(* IEC 61131-3 sources: rusty/tests/lit/single/builtin, 48 files *)

(* ---- abs_arguments.st ---- *)
// RUN: %COMPILE %s && %RUN | %CHECK %s
//
// ABS gives the same result for the implicit (positional) and the explicit (named) call form.

FUNCTION main
VAR
    neg : DINT := -42;
    a   : DINT;
    b   : DINT;
END_VAR

a := ABS(neg);
b := ABS(IN := neg);
// CHECK: ABS=42 42
printf('ABS=%d %d$N', a, b);
END_FUNCTION

(* ---- abs_floats.st ---- *)
// RUN: %COMPILE %s && %RUN | %CHECK %s
//
// ABS on floats lowers to the llvm.fabs intrinsic.

FUNCTION main

// CHECK: real=3.2 0.0 3.3 0.0
printf('real=%.1f %.1f %.1f %.1f$N', ABS(REAL#-3.2), ABS(REAL#-0.0), ABS(REAL#3.3), ABS(REAL#0.0));

// CHECK: lreal=2.5 0.0 2.6 0.0
printf('lreal=%.1f %.1f %.1f %.1f$N', ABS(LREAL#-2.5), ABS(LREAL#-0.0), ABS(LREAL#2.6), ABS(LREAL#0.0));
END_FUNCTION

(* ---- abs_signed.st ---- *)
// RUN: %COMPILE %s && %RUN | %CHECK %s
//
// ABS is a builtin; signed integers lower to the llvm.abs intrinsic with
// is_int_min_poison = false, so ABS(INT_MIN) wraps to INT_MIN.

FUNCTION main
VAR
    min : INT := INT#-32768;
END_VAR

// CHECK: sint=120 0 121 0
printf('sint=%d %d %d %d$N', ABS(SINT#-120), ABS(SINT#-0), ABS(SINT#121), ABS(SINT#0));

// CHECK: int=99 0 98 0
printf('int=%d %d %d %d$N', ABS(INT#-99), ABS(INT#-0), ABS(INT#98), ABS(INT#0));

// CHECK: dint=77 0 78 0
printf('dint=%d %d %d %d$N', ABS(-77), ABS(-0), ABS(78), ABS(0));

// CHECK: lint=88 0 89 0
printf('lint=%lld %lld %lld %lld$N', ABS(LINT#-88), ABS(LINT#-0), ABS(LINT#89), ABS(LINT#0));

// CHECK: big=1234567890123
printf('big=%lld$N', ABS(LINT#-1234567890123));

// CHECK: min=-32768
printf('min=%d$N', ABS(min));

// explicit calls to the library monomorphs still link against the stdlib
// CHECK: lib=7
printf('lib=%d$N', ABS__DINT(DINT#-7));
END_FUNCTION

(* ---- abs_unsigned.st ---- *)
// RUN: %COMPILE %s && %RUN | %CHECK %s
//
// ABS of an unsigned value returns the value unchanged instead of calling a
// non-existent monomorph (previously a crash at runtime). Each call reports
// warning E150, see abs_unsigned_warning.st.

FUNCTION main
VAR
    u8  : USINT := USINT#200;
    u16 : UINT  := UINT#5;
    u32 : UDINT := UDINT#4000000000;
    u64 : ULINT := ULINT#42;
END_VAR

// CHECK: u8=200
printf('u8=%d$N', ABS(u8));

// CHECK: u16=5
printf('u16=%d$N', ABS(u16));

// CHECK: u32=4000000000
printf('u32=%u$N', ABS(u32));

// CHECK: u64=42
printf('u64=%llu$N', ABS(u64));
END_FUNCTION

(* ---- abs_unsigned_warning.st ---- *)
// RUN: %COMPILE %s 2>&1 | %CHECK %s
//
// ABS of an unsigned value has no effect and reports a warning for each call.

FUNCTION main
VAR
    u8  : USINT;
    u16 : UINT;
    u32 : UDINT;
    u64 : ULINT;
    res : ULINT;
END_VAR

// CHECK: {{.*}}warning[E150]{{.*}}ABS on a value of unsigned type 'USINT' has no effect{{.*}}
res := ABS(u8);

// CHECK: {{.*}}warning[E150]{{.*}}ABS on a value of unsigned type 'UINT' has no effect{{.*}}
res := ABS(u16);

// CHECK: {{.*}}warning[E150]{{.*}}ABS on a value of unsigned type 'UDINT' has no effect{{.*}}
res := ABS(u32);

// CHECK: {{.*}}warning[E150]{{.*}}ABS on a value of unsigned type 'ULINT' has no effect{{.*}}
res := ABS(u64);
END_FUNCTION

(* ---- add_arguments.st ---- *)
// RUN: %COMPILE %s && %RUN | %CHECK %s
//
// ADD declares a single variadic parameter. A variadic parameter cannot be named, thus ADD has an
// implicit (positional) call form only. The form is extensible.

FUNCTION main
VAR
    x : DINT := 9;
    y : DINT := 7331;
    z : DINT := 60;
    a : DINT;
    b : DINT;
END_VAR

a := ADD(x, y);
b := ADD(x, y, z);
// CHECK: ADD=7340 7400
printf('ADD=%d %d$N', a, b);
END_FUNCTION

(* ---- add_mul_named_argument.st ---- *)
// RUN: not %COMPILE %s --error-format clang 2>&1 | %CHECK %s
//
// ADD and MUL declare a single variadic parameter, which has no name. A named argument is
// rejected, also IN1 and also with the standard library linked.

FUNCTION main : DINT
VAR
    a : DINT := 1;
    b : DINT := 2;
END_VAR
    // CHECK: {{.*}}add_mul_named_argument.st:[[@LINE+2]]:{{[0-9]+}}:{{.*}}error[E089]: Invalid call parameters
    // CHECK-NEXT: {{.*}}add_mul_named_argument.st:[[@LINE+1]]:{{[0-9]+}}:{{.*}}error[E048]: Could not resolve reference to IN1
    main := ADD(IN1 := a, b);
    // CHECK-NEXT: {{.*}}add_mul_named_argument.st:[[@LINE+2]]:{{[0-9]+}}:{{.*}}error[E089]: Invalid call parameters
    // CHECK-NEXT: {{.*}}add_mul_named_argument.st:[[@LINE+1]]:{{[0-9]+}}:{{.*}}error[E048]: Could not resolve reference to IN1
    main := MUL(IN1 := a, b);
    // CHECK-NEXT: error: Compilation aborted due to critical errors
END_FUNCTION

(* ---- adr_arguments.st ---- *)
// RUN: %COMPILE %s && %RUN | %CHECK %s
//
// ADR returns the same address for the implicit (positional) and the explicit (named) call form.

FUNCTION main
VAR
    i : INT := 5;
    p : BOOL;
END_VAR

p := ADR(i) = ADR(IN := i);
// CHECK: ADR=1
printf('ADR=%d$N', p);
END_FUNCTION

(* ---- adr_ptr_arith_runtime.st ---- *)
// RUN: %COMPILE %s && %RUN | %CHECK %s
//
// `ADR(x) + N` is byte-stride pointer arithmetic — `ADR` is declared to
// return LWORD, so the `+` flows through the integer-arithmetic path; the
// receiver pointer ends up `N` bytes past the operand. Regression for #1749
// (previously panicked in `create_llvm_int_binary_expression`).

FUNCTION main
VAR
    arr : ARRAY[0..7] OF BYTE := [0, 0, 0, 0, 0, 0, 0, 0];
    pt  : REF_TO BYTE;
END_VAR

pt := ADR(arr) + 4;
pt^ := BYTE#16#AB;

// CHECK: arr[4]=171
printf('arr[4]=%d$N', arr[4]);

pt := ADR(arr) + 7;
pt^ := BYTE#16#5C;

// CHECK: arr[7]=92
printf('arr[7]=%d$N', arr[7]);

// Subtraction flows through the same path: take a pointer past the end
// and walk back. Writing to arr[2] via `ADR(arr[6]) - 4`.
pt := ADR(arr[6]) - 4;
pt^ := BYTE#16#11;

// CHECK: arr[2]=17
printf('arr[2]=%d$N', arr[2]);
END_FUNCTION

(* ---- and_arguments.st ---- *)
// RUN: %COMPILE %s && %RUN | %CHECK %s
//
// AND declares a single variadic parameter. A variadic parameter cannot be named, thus AND has an
// implicit (positional) call form only. The form is extensible. AND gives the same result as the
// `AND` operator, for BOOL values as well as for bit and integer values.

FUNCTION main
VAR
    t : BOOL := TRUE;
    f : BOOL := FALSE;
    x : BYTE := 16#F0;
    y : BYTE := 16#3C;
    z : BYTE := 16#18;
    i : DINT := 12;
    j : DINT := 10;
    a : BOOL;
    b : BOOL;
    c : BYTE;
    d : BYTE;
    e : DINT;
END_VAR

a := AND(t, t);
b := AND(t, t, f);
// CHECK: AND=1 0 1 0
printf('AND=%u %u %u %u$N', a, b, t AND t, t AND t AND f);

c := AND(x, y);
d := AND(x, y, z);
e := AND(i, j);
// CHECK: AND-bits=48 16 8
printf('AND-bits=%u %u %d$N', c, d, e);
// CHECK: AND-bits-operator=48 16 8
printf('AND-bits-operator=%u %u %d$N', x AND y, x AND y AND z, i AND j);
END_FUNCTION

(* ---- arithmetic_bit_strings.st ---- *)
// RUN: %COMPILE %s 2> %t.err && %RUN | %CHECK %s
// RUN: not grep -E "error|warning" %t.err
//
// ADD, SUB, MUL and DIV accept bit strings as their operators do, and compute the same values.

FUNCTION main : DINT
VAR
    b : BYTE := 16#FF;
    dw : DWORD := 16#100;
    di : DINT := 7;
END_VAR

// CHECK: ADD BYTE 256 256
printf('ADD BYTE %u %u$N', ADD(b, 1), b + 1);
// CHECK-NEXT: SUB DWORD 255 255
printf('SUB DWORD %u %u$N', SUB(dw, 1), dw - 1);
// CHECK-NEXT: SUB named 255 255
printf('SUB named %u %u$N', SUB(IN2 := 1, IN1 := dw), dw - 1);
// CHECK-NEXT: MUL DWORD 65536 65536
printf('MUL DWORD %u %u$N', MUL(dw, dw), dw * dw);
// CHECK-NEXT: DIV DWORD 128 128
printf('DIV DWORD %u %u$N', DIV(dw, 2), dw / 2);
// CHECK-NEXT: ADD DINT BYTE 262 262
printf('ADD DINT BYTE %d %d$N', ADD(di, b), di + b);
END_FUNCTION

(* ---- datetime_arithmetic_chain.st ---- *)
// RUN: %COMPILE %s && %RUN | %CHECK %s
// Chains of date and time arithmetic, in operator and builtin form

FUNCTION main
    VAR
        x : DT := DT#2027-05-05-22:30:15;
        y : TIME := TIME#20s;
        z : TOD := TOD#23:58:00;
    END_VAR

    x := x + y + y + TIME#2h555s;
    printf('%s$N', REF(DT_TO_STRING(x)));                                           // CHECK: DT#2027-05-06-00:40:10

    z := z + TIME#2m5s;
    printf('%s$N', REF(TOD_TO_STRING(z)));                                          // CHECK: TOD#00:00:05

    x := ADD(x, y, MUL(y, 2));
    printf('%s$N', REF(DT_TO_STRING(x)));                                           // CHECK: DT#2027-05-06-00:41:10

    z := SUB(z, TIME#10s);
    printf('%s$N', REF(TOD_TO_STRING(z)));                                          // CHECK: TOD#23:59:55

END_FUNCTION

(* ---- datetime_arithmetic_date.st ---- *)
// RUN: %COMPILE %s && %RUN | %CHECK %s
// Test DATE arithmetic operations return correct types and values

FUNCTION main
    VAR
        date1 : DATE;
        date2 : DATE;
        result : TIME;
    END_VAR

    // SUB_DATE_DATE: DATE - DATE -> TIME (u32)
    date1 := DATE#2024-01-15;
    date2 := DATE#2024-01-10;
    result := SUB_DATE_DATE(date1, date2);
    printf('%s$N', REF(TIME_TO_STRING(result)));                                    // CHECK: T#5d

    // The operators carry out the same functions
    result := date1 - date2;
    printf('%s$N', REF(TIME_TO_STRING(result)));                                    // CHECK: T#5d

    // The builtins carry out the same functions as the operators
    result := SUB(date1, date2);
    printf('%s$N', REF(TIME_TO_STRING(result)));                                    // CHECK: T#5d

END_FUNCTION

(* ---- datetime_arithmetic_dt.st ---- *)
// RUN: %COMPILE %s && %RUN | %CHECK %s
// Test DT arithmetic operations return correct types and values

FUNCTION main
    VAR
        dt1 : DT;
        dt2 : DT;
        t1 : TIME;
        result : TIME;
        dt_result : DT;
    END_VAR

    // ADD_DT_TIME: DT + TIME -> DT (u32)
    dt1 := DT#2024-01-15-12:30:00;
    t1 := TIME#5s;
    dt_result := ADD_DT_TIME(dt1, t1);
    printf('%s$N', REF(DT_TO_STRING(dt_result)));                                   // CHECK: DT#2024-01-15-12:30:05

    // SUB_DT_TIME: DT - TIME -> DT (u32)
    dt1 := DT#2024-01-15-12:30:05;
    t1 := TIME#3s;
    dt_result := SUB_DT_TIME(dt1, t1);
    printf('%s$N', REF(DT_TO_STRING(dt_result)));                                   // CHECK: DT#2024-01-15-12:30:02

    // SUB_DT_DT: DT - DT -> TIME (u32)
    dt1 := DT#2024-01-15-12:30:10;
    dt2 := DT#2024-01-15-12:30:00;
    result := SUB_DT_DT(dt1, dt2);
    printf('%s$N', REF(TIME_TO_STRING(result)));                                    // CHECK: T#10s

    // The operators carry out the same functions
    dt_result := dt1 + t1;
    printf('%s$N', REF(DT_TO_STRING(dt_result)));                                   // CHECK: DT#2024-01-15-12:30:13
    dt_result := dt1 - t1;
    printf('%s$N', REF(DT_TO_STRING(dt_result)));                                   // CHECK: DT#2024-01-15-12:30:07
    result := dt1 - dt2;
    printf('%s$N', REF(TIME_TO_STRING(result)));                                    // CHECK: T#10s

    // The builtins carry out the same functions as the operators
    dt_result := ADD(dt1, t1, T#1m);
    printf('%s$N', REF(DT_TO_STRING(dt_result)));                                   // CHECK: DT#2024-01-15-12:31:13
    result := SUB(dt1, dt2);
    printf('%s$N', REF(TIME_TO_STRING(result)));                                    // CHECK: T#10s

END_FUNCTION

(* ---- datetime_arithmetic_ldate.st ---- *)
// RUN: %COMPILE %s && %RUN | %CHECK %s
// Test LDATE arithmetic operations return correct types and values

FUNCTION main
    VAR
        ldate1 : LDATE;
        ldate2 : LDATE;
        lresult : LTIME;
    END_VAR

    // SUB_LDATE_LDATE: LDATE - LDATE -> LTIME (i64)
    ldate1 := LDATE#2024-01-15;
    ldate2 := LDATE#2024-01-10;
    lresult := SUB_LDATE_LDATE(ldate1, ldate2);
    printf('%s$N', REF(LTIME_TO_STRING(lresult)));                                  // CHECK: LTIME#5d

    // The operators carry out the same functions
    lresult := ldate1 - ldate2;
    printf('%s$N', REF(LTIME_TO_STRING(lresult)));                                  // CHECK: LTIME#5d

    // The builtins carry out the same functions as the operators
    lresult := SUB(ldate1, ldate2);
    printf('%s$N', REF(LTIME_TO_STRING(lresult)));                                  // CHECK: LTIME#5d

END_FUNCTION

(* ---- datetime_arithmetic_ldt.st ---- *)
// RUN: %COMPILE %s && %RUN | %CHECK %s
// Test LDT arithmetic operations return correct types and values

FUNCTION main
    VAR
        ldt1 : LDT;
        ldt2 : LDT;
        lt1 : LTIME;
        lresult : LTIME;
        ldt_result : LDT;
    END_VAR

    // ADD_LDT_LTIME: LDT + LTIME -> LDT (i64, nanosecond precision)
    ldt1 := LDT#2024-01-15-12:30:00;
    lt1 := LTIME#5s;
    ldt_result := ADD_LDT_LTIME(ldt1, lt1);
    printf('%s$N', REF(LDT_TO_STRING(ldt_result)));                                 // CHECK: LDT#2024-01-15-12:30:05

    // SUB_LDT_LTIME: LDT - LTIME -> LDT (i64)
    ldt1 := LDT#2024-01-15-12:30:05;
    lt1 := LTIME#3s;
    ldt_result := SUB_LDT_LTIME(ldt1, lt1);
    printf('%s$N', REF(LDT_TO_STRING(ldt_result)));                                 // CHECK: LDT#2024-01-15-12:30:02

    // SUB_LDT_LDT: LDT - LDT -> LTIME (i64, result is difference in nanoseconds)
    ldt1 := LDT#2024-01-15-12:30:10;
    ldt2 := LDT#2024-01-15-12:30:00;
    lresult := SUB_LDT_LDT(ldt1, ldt2);
    printf('%s$N', REF(LTIME_TO_STRING(lresult)));                                  // CHECK: LTIME#10s

    // The operators carry out the same functions
    ldt_result := ldt1 + lt1;
    printf('%s$N', REF(LDT_TO_STRING(ldt_result)));                                 // CHECK: LDT#2024-01-15-12:30:13
    ldt_result := ldt1 - lt1;
    printf('%s$N', REF(LDT_TO_STRING(ldt_result)));                                 // CHECK: LDT#2024-01-15-12:30:07
    lresult := ldt1 - ldt2;
    printf('%s$N', REF(LTIME_TO_STRING(lresult)));                                  // CHECK: LTIME#10s

    // The builtins carry out the same functions as the operators
    ldt_result := ADD(ldt1, lt1, lt1);
    printf('%s$N', REF(LDT_TO_STRING(ldt_result)));                                 // CHECK: LDT#2024-01-15-12:30:16
    lresult := SUB(ldt1, ldt2);
    printf('%s$N', REF(LTIME_TO_STRING(lresult)));                                  // CHECK: LTIME#10s

END_FUNCTION

(* ---- datetime_arithmetic_long_chain.st ---- *)
// RUN: %COMPILE %s && %RUN | %CHECK %s
// A long chain of date and time arithmetic compiles in time linear to its length

FUNCTION main
    VAR
        t : TIME := TIME#1s;
    END_VAR

    t := ADD(t, t, t, t, t, t, t, t, t, t, t, t, t, t, t, t, t, t, t, t, t, t, t, t, t, t, t, t, t, t);
    printf('%s$N', REF(TIME_TO_STRING(t)));                                         // CHECK: T#30s

    t := t + t + t + t + t + t + t + t + t + t + t + t + t + t + t + t + t + t + t + t + t + t + t + t + t + t + t + t + t + t;
    printf('%s$N', REF(TIME_TO_STRING(t)));                                         // CHECK: T#15m

END_FUNCTION

(* ---- datetime_arithmetic_ltime.st ---- *)
// RUN: %COMPILE %s && %RUN | %CHECK %s
// Test LTIME arithmetic operations return correct types and values

FUNCTION main
    VAR
        lt1 : LTIME;
        lt2 : LTIME;
        lresult : LTIME;
    END_VAR

    // ADD_LTIME: LTIME + LTIME -> LTIME (i64)
    lt1 := LTIME#5s;
    lt2 := LTIME#3s;
    lresult := ADD_LTIME(lt1, lt2);
    printf('%s$N', REF(LTIME_TO_STRING(lresult)));                                  // CHECK: LTIME#8s

    // SUB_LTIME: LTIME - LTIME -> LTIME (i64)
    lt1 := LTIME#10s;
    lt2 := LTIME#3s;
    lresult := SUB_LTIME(lt1, lt2);
    printf('%s$N', REF(LTIME_TO_STRING(lresult)));                                  // CHECK: LTIME#7s

    // The operators carry out the same functions
    lresult := lt1 + lt2;
    printf('%s$N', REF(LTIME_TO_STRING(lresult)));                                  // CHECK: LTIME#13s
    lresult := lt1 - lt2;
    printf('%s$N', REF(LTIME_TO_STRING(lresult)));                                  // CHECK: LTIME#7s
    lresult := lt1 * 2;
    printf('%s$N', REF(LTIME_TO_STRING(lresult)));                                  // CHECK: LTIME#20s
    lresult := 2 * lt1;
    printf('%s$N', REF(LTIME_TO_STRING(lresult)));                                  // CHECK: LTIME#20s
    lresult := lt1 / 4;
    printf('%s$N', REF(LTIME_TO_STRING(lresult)));                                  // CHECK: LTIME#2s500ms

    // The builtins carry out the same functions as the operators
    lresult := ADD(lt1, lt2, LTIME#1s);
    printf('%s$N', REF(LTIME_TO_STRING(lresult)));                                  // CHECK: LTIME#14s
    lresult := MUL(lt1, 1.5);
    printf('%s$N', REF(LTIME_TO_STRING(lresult)));                                  // CHECK: LTIME#15s

END_FUNCTION

(* ---- datetime_arithmetic_ltod.st ---- *)
// RUN: %COMPILE %s && %RUN | %CHECK %s
// Test LTOD arithmetic operations return correct types and values

FUNCTION main
    VAR
        ltod1 : LTOD;
        ltod2 : LTOD;
        lt1 : LTIME;
        lresult : LTIME;
        ltod_result : LTOD;
    END_VAR

    // ADD_LTOD_LTIME: LTOD + LTIME -> LTOD (wraps at day boundary)
    ltod1 := LTOD#23:59:50;
    lt1 := LTIME#20s;
    ltod_result := ADD_LTOD_LTIME(ltod1, lt1);
    printf('%s$N', REF(LTOD_TO_STRING(ltod_result)));                               // CHECK: LTOD#00:00:10

    // SUB_LTOD_LTIME: LTOD - LTIME -> LTOD
    ltod1 := LTOD#00:01:00;
    lt1 := LTIME#30s;
    ltod_result := SUB_LTOD_LTIME(ltod1, lt1);
    printf('%s$N', REF(LTOD_TO_STRING(ltod_result)));                               // CHECK: LTOD#00:00:30

    // SUB_LTOD_LTOD: LTOD - LTOD -> LTIME (i64)
    ltod1 := LTOD#10:30:00;
    ltod2 := LTOD#10:20:00;
    lresult := SUB_LTOD_LTOD(ltod1, ltod2);
    printf('%s$N', REF(LTIME_TO_STRING(lresult)));                                  // CHECK: LTIME#10m

    // The operators carry out the same functions
    ltod_result := ltod1 + lt1;
    printf('%s$N', REF(LTOD_TO_STRING(ltod_result)));                               // CHECK: LTOD#10:30:30
    ltod_result := ltod1 - lt1;
    printf('%s$N', REF(LTOD_TO_STRING(ltod_result)));                               // CHECK: LTOD#10:29:30
    lresult := ltod1 - ltod2;
    printf('%s$N', REF(LTIME_TO_STRING(lresult)));                                  // CHECK: LTIME#10m
    ltod_result := LTOD#23:59:50 + LTIME#20s;
    printf('%s$N', REF(LTOD_TO_STRING(ltod_result)));                               // CHECK: LTOD#00:00:10

    // The builtins carry out the same functions as the operators
    ltod_result := ADD(ltod1, lt1, lt1);
    printf('%s$N', REF(LTOD_TO_STRING(ltod_result)));                               // CHECK: LTOD#10:31:00
    lresult := SUB(ltod1, ltod2);
    printf('%s$N', REF(LTIME_TO_STRING(lresult)));                                  // CHECK: LTIME#10m

END_FUNCTION

(* ---- datetime_arithmetic_time.st ---- *)
// RUN: %COMPILE %s && %RUN | %CHECK %s
// Test TIME arithmetic operations return correct types and values

FUNCTION main
    VAR
        t1 : TIME;
        t2 : TIME;
        result : TIME;
    END_VAR

    // ADD_TIME: TIME + TIME -> TIME (u32)
    t1 := TIME#5s;
    t2 := TIME#3s;
    result := ADD_TIME(t1, t2);
    printf('%s$N', REF(TIME_TO_STRING(result)));                                    // CHECK: T#8s

    // SUB_TIME: TIME - TIME -> TIME (u32)
    t1 := TIME#10s;
    t2 := TIME#3s;
    result := SUB_TIME(t1, t2);
    printf('%s$N', REF(TIME_TO_STRING(result)));                                    // CHECK: T#7s

    // The operators carry out the same functions
    result := t1 + t2;
    printf('%s$N', REF(TIME_TO_STRING(result)));                                    // CHECK: T#13s
    result := t1 - t2;
    printf('%s$N', REF(TIME_TO_STRING(result)));                                    // CHECK: T#7s
    result := t1 * 3;
    printf('%s$N', REF(TIME_TO_STRING(result)));                                    // CHECK: T#30s
    result := 2 * t1;
    printf('%s$N', REF(TIME_TO_STRING(result)));                                    // CHECK: T#20s
    result := t1 / 4;
    printf('%s$N', REF(TIME_TO_STRING(result)));                                    // CHECK: T#2s500ms
    result := t1 + 5;
    printf('%s$N', REF(TIME_TO_STRING(result)));                                    // CHECK: T#10s5ms

    // The builtins carry out the same functions as the operators
    result := ADD(t1, t2, T#1s);
    printf('%s$N', REF(TIME_TO_STRING(result)));                                    // CHECK: T#14s
    result := SUB(t1, t2);
    printf('%s$N', REF(TIME_TO_STRING(result)));                                    // CHECK: T#7s
    result := MUL(t1, 1.5);
    printf('%s$N', REF(TIME_TO_STRING(result)));                                    // CHECK: T#15s
    result := DIV(t1, 2.5);
    printf('%s$N', REF(TIME_TO_STRING(result)));                                    // CHECK: T#4s

END_FUNCTION

(* ---- datetime_arithmetic_tod.st ---- *)
// RUN: %COMPILE %s && %RUN | %CHECK %s
// Test TOD arithmetic operations return correct types and values

FUNCTION main
    VAR
        tod1 : TOD;
        tod2 : TOD;
        t1 : TIME;
        result : TIME;
        tod_result : TOD;
    END_VAR

    // ADD_TOD_TIME: TOD + TIME -> TOD (wraps at day boundary)
    tod1 := TOD#23:59:50;
    t1 := TIME#20s;
    result := ADD_TOD_TIME(tod1, t1);
    printf('%s$N', REF(TOD_TO_STRING(result)));                                     // CHECK: TOD#00:00:10

    // SUB_TOD_TIME: TOD - TIME -> TOD
    tod1 := TOD#00:01:00;
    t1 := TIME#30s;
    result := SUB_TOD_TIME(tod1, t1);
    printf('%s$N', REF(TOD_TO_STRING(result)));                                     // CHECK: TOD#00:00:30

    // SUB_TOD_TOD: TOD - TOD -> TIME (u32)
    tod1 := TOD#10:30:00;
    tod2 := TOD#10:20:00;
    result := SUB_TOD_TOD(tod1, tod2);
    printf('%s$N', REF(TIME_TO_STRING(result)));                                    // CHECK: T#10m

    // Test ADD_TOD_TIME with simple arithmetic
    tod1 := TOD#12:00:00;
    t1 := TIME#1m;
    result := ADD_TOD_TIME(tod1, t1);
    printf('%s$N', REF(TOD_TO_STRING(result)));                                     // CHECK: TOD#12:01:00

    // Test SUB_TOD_TIME with simple case
    tod1 := TOD#12:05:00;
    t1 := TIME#1m;
    result := SUB_TOD_TIME(tod1, t1);
    printf('%s$N', REF(TOD_TO_STRING(result)));                                     // CHECK: TOD#12:04:00

    // The operators carry out the same functions
    tod_result := tod1 + t1;
    printf('%s$N', REF(TOD_TO_STRING(tod_result)));                                 // CHECK: TOD#12:06:00
    tod_result := tod1 - t1;
    printf('%s$N', REF(TOD_TO_STRING(tod_result)));                                 // CHECK: TOD#12:04:00
    result := tod1 - tod2;
    printf('%s$N', REF(TIME_TO_STRING(result)));                                    // CHECK: T#1h45m
    tod_result := TOD#23:59:50 + TIME#20s;
    printf('%s$N', REF(TOD_TO_STRING(tod_result)));                                 // CHECK: TOD#00:00:10

    // The builtins carry out the same functions as the operators
    tod_result := ADD(tod1, t1, TIME#20s);
    printf('%s$N', REF(TOD_TO_STRING(tod_result)));                                 // CHECK: TOD#12:06:20
    tod_result := SUB(tod1, t1);
    printf('%s$N', REF(TOD_TO_STRING(tod_result)));                                 // CHECK: TOD#12:04:00
    result := SUB(tod1, tod2);
    printf('%s$N', REF(TIME_TO_STRING(result)));                                    // CHECK: T#1h45m

END_FUNCTION

(* ---- div_arguments.st ---- *)
// RUN: %COMPILE %s && %RUN | %CHECK %s
//
// DIV gives the same result for the implicit (positional) and the explicit (named) call form, in
// declaration order and reordered. A call may also mix both forms: a named argument claims the slot
// its name declares, and the positional arguments fill the remaining slots in the order they are
// written.

FUNCTION main
VAR
    x : DINT := 9;
    y : DINT := 7331;
    a : DINT;
    b : DINT;
    c : DINT;
END_VAR

a := DIV(y, x);
b := DIV(IN1 := y, IN2 := x);
c := DIV(IN2 := x, IN1 := y);
// CHECK: DIV=814 814 814
printf('DIV=%d %d %d$N', a, b, c);

// named argument before the positional one, IN1 is filled by y
a := DIV(IN2 := x, y);
// CHECK: DIV-named-first=814
printf('DIV-named-first=%d$N', a);
END_FUNCTION

(* ---- eq_arguments.st ---- *)
// RUN: %COMPILE %s && %RUN | %CHECK %s
//
// EQ declares a single variadic parameter. A variadic parameter cannot be named, thus EQ has an
// implicit (positional) call form only. The form is extensible: every neighbouring pair is compared
// and the results are combined with AND.

FUNCTION main
VAR
    a : DINT := 30;
    b : DINT := 20;
    c : DINT := 10;
    p : BOOL;
    q : BOOL;
    r : BOOL;
END_VAR

p := EQ(b, b);
q := EQ(b, b, b);
r := EQ(a, b, b);
// CHECK: EQ=1 1 0
printf('EQ=%d %d %d$N', p, q, r);
END_FUNCTION

(* ---- function_named_like_builtin.st ---- *)
// RUN: not %COMPILE %s --error-format clang 2>&1 | %CHECK %s
// A POU that takes the name of a built-in function is rejected with a message that names the collision.

// CHECK: {{.*}}error[E004]: `ABS` is the name of a built-in function
FUNCTION ABS : DINT
VAR_INPUT
    IN : DINT;
END_VAR
END_FUNCTION

// CHECK-NEXT: {{.*}}error[E004]: `Sel` is the name of a built-in function
FUNCTION Sel : DINT
VAR_INPUT
    G : BOOL;
    IN0 : DINT;
    IN1 : DINT;
END_VAR
END_FUNCTION

// CHECK-NEXT: error: Compilation aborted due to critical errors

(* ---- ge_arguments.st ---- *)
// RUN: %COMPILE %s && %RUN | %CHECK %s
//
// GE declares a single variadic parameter. A variadic parameter cannot be named, thus GE has an
// implicit (positional) call form only. The form is extensible: every neighbouring pair is compared
// and the results are combined with AND.

FUNCTION main
VAR
    a : DINT := 30;
    b : DINT := 20;
    c : DINT := 10;
    p : BOOL;
    q : BOOL;
    r : BOOL;
END_VAR

p := GE(a, b);
q := GE(a, b, c);
r := GE(a, c, b);
// CHECK: GE=1 1 0
printf('GE=%d %d %d$N', p, q, r);
END_FUNCTION

(* ---- gt_arguments.st ---- *)
// RUN: %COMPILE %s && %RUN | %CHECK %s
//
// GT declares a single variadic parameter. A variadic parameter cannot be named, thus GT has an
// implicit (positional) call form only. The form is extensible: every neighbouring pair is compared
// and the results are combined with AND.

FUNCTION main
VAR
    a : DINT := 30;
    b : DINT := 20;
    c : DINT := 10;
    p : BOOL;
    q : BOOL;
    r : BOOL;
END_VAR

p := GT(a, b);
q := GT(a, b, c);
r := GT(a, c, b);
// CHECK: GT=1 1 0
printf('GT=%d %d %d$N', p, q, r);
END_FUNCTION

(* ---- le_arguments.st ---- *)
// RUN: %COMPILE %s && %RUN | %CHECK %s
//
// LE declares a single variadic parameter. A variadic parameter cannot be named, thus LE has an
// implicit (positional) call form only. The form is extensible: every neighbouring pair is compared
// and the results are combined with AND.

FUNCTION main
VAR
    a : DINT := 30;
    b : DINT := 20;
    c : DINT := 10;
    p : BOOL;
    q : BOOL;
    r : BOOL;
END_VAR

p := LE(c, b);
q := LE(c, b, a);
r := LE(c, a, b);
// CHECK: LE=1 1 0
printf('LE=%d %d %d$N', p, q, r);
END_FUNCTION

(* ---- lower_bound_arguments.st ---- *)
// RUN: %COMPILE %s && %RUN | %CHECK %s
//
// LOWER_BOUND gives the same result for the implicit (positional) and the explicit (named) call form,
// in declaration order and reordered.

FUNCTION main
VAR
    arr : ARRAY[0..9] OF BYTE := [0, 1, 2, 3, 4, 5, 6, 7, 8, 9];
END_VAR

bounds(arr);
END_FUNCTION

FUNCTION bounds : DINT
VAR_IN_OUT
    vla : ARRAY[*] OF BYTE;
END_VAR
VAR
    dim : DINT := 1;
    a   : DINT;
    b   : DINT;
    c   : DINT;
END_VAR

a := LOWER_BOUND(vla, dim);
b := LOWER_BOUND(ARR := vla, DIM := dim);
c := LOWER_BOUND(DIM := dim, ARR := vla);
// CHECK: LOWER_BOUND=0 0 0
printf('LOWER_BOUND=%d %d %d$N', a, b, c);
END_FUNCTION

(* ---- lt_arguments.st ---- *)
// RUN: %COMPILE %s && %RUN | %CHECK %s
//
// LT declares a single variadic parameter. A variadic parameter cannot be named, thus LT has an
// implicit (positional) call form only. The form is extensible: every neighbouring pair is compared
// and the results are combined with AND.

FUNCTION main
VAR
    a : DINT := 30;
    b : DINT := 20;
    c : DINT := 10;
    p : BOOL;
    q : BOOL;
    r : BOOL;
END_VAR

p := LT(c, b);
q := LT(c, b, a);
r := LT(c, a, b);
// CHECK: LT=1 1 0
printf('LT=%d %d %d$N', p, q, r);
END_FUNCTION

(* ---- mod_arguments.st ---- *)
// RUN: %COMPILE %s && %RUN | %CHECK %s
//
// MOD gives the same result for the implicit (positional) and the explicit (named) call form, in
// declaration order and reordered. MOD gives the same result as the `MOD` operator, for integer as
// well as for REAL values, and for two TIME or two LTIME values.

FUNCTION main
VAR
    x : DINT := 9;
    y : DINT := 7331;
    a : DINT;
    b : DINT;
    c : DINT;
    r : REAL := 7.5;
    s : REAL := 2.0;
    q : REAL;
    t1 : TIME := T#7s;
    t2 : TIME := T#3s;
    t : TIME;
    lt1 : LTIME := LTIME#7s500ms;
    lt2 : LTIME := LTIME#2s;
    lt : LTIME;
END_VAR

a := MOD(y, x);
b := MOD(IN1 := y, IN2 := x);
c := MOD(IN2 := x, IN1 := y);
// CHECK: MOD=5 5 5 5
printf('MOD=%d %d %d %d$N', a, b, c, y MOD x);

q := MOD(r, s);
// CHECK: MOD-real=1.5 1.5
printf('MOD-real=%.1f %.1f$N', q, r MOD s);

t := MOD(t1, t2);
// CHECK: MOD-time=T#1s
printf('MOD-time=%s$N', REF(TIME_TO_STRING(t)));

lt := MOD(IN2 := lt2, IN1 := lt1);
// CHECK: MOD-ltime=LTIME#1s500ms
printf('MOD-ltime=%s$N', REF(LTIME_TO_STRING(lt)));
END_FUNCTION

(* ---- move_arguments.st ---- *)
// RUN: %COMPILE %s && %RUN | %CHECK %s
//
// MOVE gives the same result for the implicit (positional) and the explicit (named) call form.

FUNCTION main
VAR
    y : DINT := 7331;
    a : DINT;
    b : DINT;
END_VAR

a := MOVE(y);
b := MOVE(IN := y);
// CHECK: MOVE=7331 7331
printf('MOVE=%d %d$N', a, b);
END_FUNCTION

(* ---- mul_arguments.st ---- *)
// RUN: %COMPILE %s && %RUN | %CHECK %s
//
// MUL declares a single variadic parameter. A variadic parameter cannot be named, thus MUL has an
// implicit (positional) call form only. The form is extensible.

FUNCTION main
VAR
    x : DINT := 9;
    a : DINT;
    b : DINT;
END_VAR

a := MUL(x, 3);
b := MUL(x, 3, 2);
// CHECK: MUL=27 54
printf('MUL=%d %d$N', a, b);
END_FUNCTION

(* ---- mux_arguments.st ---- *)
// RUN: %COMPILE %s && %RUN | %CHECK %s
//
// MUX names its first parameter K and takes the remaining ones through a variadic parameter. A
// variadic parameter cannot be named, thus only K has an explicit (named) call form.

FUNCTION main
VAR
    x : DINT := 9;
    y : DINT := 7331;
    z : DINT := 42;
    n : DINT := -1;
    a : DINT;
    b : DINT;
    c : DINT;
    lr : LREAL;
END_VAR

a := MUX(1, x, y);
b := MUX(K := 1, x, y);
// CHECK: MUX=7331 7331
printf('MUX=%d %d$N', a, b);

c := MUX(2, x, y, z);
// CHECK: MUX-extended=42
printf('MUX-extended=%d$N', c);

// the variadic arguments resolve the generic type of the mixed call as they do in the positional call,
// thus a negative value keeps its sign when it is widened
lr := MUX(0, n, x);
// CHECK: MUX-widened=-1.0
printf('MUX-widened=%.1f$N', lr);
lr := MUX(K := 0, n, x);
// CHECK: MUX-mixed-widened=-1.0
printf('MUX-mixed-widened=%.1f$N', lr);
END_FUNCTION

(* ---- ne_arguments.st ---- *)
// RUN: %COMPILE %s && %RUN | %CHECK %s
//
// NE gives the same result for the implicit (positional) and the explicit (named) call form, in
// declaration order and reordered. A call may also mix both forms: a named argument claims the slot
// its name declares, and the positional arguments fill the remaining slots in the order they are
// written.

FUNCTION main
VAR
    lr : LREAL := 1.5;
    x  : DINT  := 9;
    y  : DINT  := 7331;
    p  : BOOL;
    q  : BOOL;
    r  : BOOL;
END_VAR

p := NE(lr, 0);
q := NE(IN1 := lr, IN2 := 0);
r := NE(IN2 := 0, IN1 := lr);
// CHECK: NE=1 1 1
printf('NE=%d %d %d$N', p, q, r);

// a mix of implicit and explicit arguments
p := NE(lr, IN2 := 0);
q := NE(IN2 := 0, lr);
// CHECK: NE-mixed=1 1
printf('NE-mixed=%d %d$N', p, q);

// parenthesized arguments
p := NE((lr), 0);
q := NE(IN1 := (lr), IN2 := 0);
// CHECK: NE-paren=1 1
printf('NE-paren=%d %d$N', p, q);

// arguments of the same type
p := NE(x, y);
q := NE(x, x);
// CHECK: NE-same-type=1 0
printf('NE-same-type=%d %d$N', p, q);
END_FUNCTION

(* ---- not_arguments.st ---- *)
// RUN: %COMPILE %s && %RUN | %CHECK %s
//
// NOT gives the same result for the implicit (positional) and the explicit (named) call form. NOT
// gives the same result as the `NOT` operator, for BOOL values as well as for bit and integer values.

FUNCTION main
VAR
    t : BOOL := TRUE;
    x : BYTE := 16#F0;
    i : DINT := 12;
    a : BOOL;
    b : BOOL;
    c : BYTE;
    d : BYTE;
    e : DINT;
END_VAR

a := NOT(t);
b := NOT(IN := t);
// CHECK: NOT=0 0 0
printf('NOT=%u %u %u$N', a, b, NOT t);

c := NOT(x);
d := NOT(IN := x);
e := NOT(IN := i);
// CHECK: NOT-bits=15 15 -13
printf('NOT-bits=%u %u %d$N', c, d, e);
// CHECK: NOT-bits-operator=15 -13
printf('NOT-bits-operator=%u %d$N', NOT x, NOT i);
END_FUNCTION

(* ---- or_arguments.st ---- *)
// RUN: %COMPILE %s && %RUN | %CHECK %s
//
// OR declares a single variadic parameter. A variadic parameter cannot be named, thus OR has an
// implicit (positional) call form only. The form is extensible. OR gives the same result as the
// `OR` operator, for BOOL values as well as for bit and integer values.

FUNCTION main
VAR
    t : BOOL := TRUE;
    f : BOOL := FALSE;
    x : BYTE := 16#F0;
    y : BYTE := 16#0C;
    z : BYTE := 16#01;
    i : DINT := 12;
    j : DINT := 10;
    a : BOOL;
    b : BOOL;
    c : BYTE;
    d : BYTE;
    e : DINT;
END_VAR

a := OR(f, f);
b := OR(f, f, t);
// CHECK: OR=0 1 0 1
printf('OR=%u %u %u %u$N', a, b, f OR f, f OR f OR t);

c := OR(x, y);
d := OR(x, y, z);
e := OR(i, j);
// CHECK: OR-bits=252 253 14
printf('OR-bits=%u %u %d$N', c, d, e);
// CHECK: OR-bits-operator=252 253 14
printf('OR-bits-operator=%u %u %d$N', x OR y, x OR y OR z, i OR j);
END_FUNCTION

(* ---- ref_arguments.st ---- *)
// RUN: %COMPILE %s && %RUN | %CHECK %s
//
// REF returns the same pointer for the implicit (positional) and the explicit (named) call form.

FUNCTION main
VAR
    i     : INT := 5;
    ptr_a : REF_TO INT;
    ptr_b : REF_TO INT;
    p     : BOOL;
END_VAR

ptr_a := REF(i);
ptr_b := REF(IN := i);
p := ptr_a = ptr_b;
// CHECK: REF=1
printf('REF=%d$N', p);
END_FUNCTION

(* ---- sel_arguments.st ---- *)
// RUN: %COMPILE %s && %RUN | %CHECK %s
//
// SEL gives the same result for the implicit (positional) and the explicit (named) call form, in
// declaration order and reordered. A call may also mix both forms: a named argument claims the slot
// its name declares, and the positional arguments fill the remaining slots in the order they are
// written.

FUNCTION main
VAR
    x : DINT := 9;
    y : DINT := 7331;
    a : DINT;
    b : DINT;
    c : DINT;
    r0 : REAL := 1.5;
    r1 : REAL := 2.5;
    r : REAL;
    s : REAL;
END_VAR

a := SEL(TRUE, x, y);
b := SEL(G := TRUE, IN0 := x, IN1 := y);
c := SEL(IN1 := y, IN0 := x, G := TRUE);
// CHECK: SEL=7331 7331 7331
printf('SEL=%d %d %d$N', a, b, c);

// named argument before the positional ones, G and IN0 are filled by FALSE and x
a := SEL(IN1 := y, FALSE, x);
// CHECK: SEL-mixed=9
printf('SEL-mixed=%d$N', a);

// the selector G stays a BOOL when the selected type is not an integer
r := SEL(IN1 := r1, FALSE, r0);
s := SEL(IN1 := r1, TRUE, r0);
// CHECK: SEL-mixed-real=1.5 2.5
printf('SEL-mixed-real=%.1f %.1f$N', r, s);
END_FUNCTION

(* ---- shl_and_shr_must_cast_left_and_right_correctly.st ---- *)
// RUN: %COMPILE %s && %RUN | %CHECK %s

// SHL and SHR must cast left and right correctly
FUNCTION main
VAR
    value : BYTE;
END_VAR

value := BIT_LOAD_B2(BYTE#255, TRUE, 2, 2);

// CHECK: 255
printf('%d$N', value);

value := BIT_LOAD_B2(BYTE#255, FALSE, 2, 2);

// CHECK: 243
printf('%d$N', value);

END_FUNCTION

FUNCTION BIT_LOAD_B2 : BYTE
VAR_INPUT
	I : BYTE;
	D : BOOL;
	P : INT;
	N : INT;
END_VAR
VAR
    result : BYTE;
END_VAR

IF D THEN
	BIT_LOAD_B2 := ROL(SHR(BYTE#255, 8 - N) OR ROR(I, P), P);
ELSE
	BIT_LOAD_B2 := ROL(SHL(BYTE#255, N) AND ROR(I, P), P);
END_IF;

END_FUNCTION

(* ---- shl_arguments.st ---- *)
// RUN: %COMPILE %s && %RUN | %CHECK %s
//
// SHL gives the same result for the implicit (positional) and the explicit (named) call form, in
// declaration order and reordered. A call may also mix both forms: a named argument claims the slot
// its name declares, and the positional arguments fill the remaining slots in the order they are
// written.

FUNCTION main
VAR
    x : DINT := 9;
    a : DINT;
    b : DINT;
    c : DINT;
END_VAR

a := SHL(x, 2);
b := SHL(IN := x, N := 2);
c := SHL(N := 2, IN := x);
// CHECK: SHL=36 36 36
printf('SHL=%d %d %d$N', a, b, c);

// named argument before the positional one, IN is filled by x
a := SHL(N := 2, x);
// CHECK: SHL-named-first=36
printf('SHL-named-first=%d$N', a);
END_FUNCTION

(* ---- shl_must_be_usable_with_integers.st ---- *)
// RUN: %COMPILE %s && %RUN | %CHECK %s

// SHL must be usable with integers
FUNCTION main
VAR
    a : INT;
END_VAR
a := SHL(21,2);

// CHECK: 84
printf('%d$N', a);
END_FUNCTION

(* ---- shr_arguments.st ---- *)
// RUN: %COMPILE %s && %RUN | %CHECK %s
//
// SHR gives the same result for the implicit (positional) and the explicit (named) call form, in
// declaration order and reordered. A call may also mix both forms: a named argument claims the slot
// its name declares, and the positional arguments fill the remaining slots in the order they are
// written.

FUNCTION main
VAR
    x : DINT := 9;
    a : DINT;
    b : DINT;
    c : DINT;
END_VAR

a := SHR(x, 2);
b := SHR(IN := x, N := 2);
c := SHR(N := 2, IN := x);
// CHECK: SHR=2 2 2
printf('SHR=%d %d %d$N', a, b, c);

// named argument before the positional one, IN is filled by x
a := SHR(N := 2, x);
// CHECK: SHR-named-first=2
printf('SHR-named-first=%d$N', a);
END_FUNCTION

(* ---- shr_must_be_usable_with_integers.st ---- *)
// RUN: %COMPILE %s && %RUN | %CHECK %s

// SHR must be usable with integers
FUNCTION main
VAR
    a : INT;
END_VAR
a := SHR(21,2);

// CHECK: 5
printf('%d$N', a);
END_FUNCTION

(* ---- shr_unsigned_byte_logical_shift.st ---- *)
// RUN: %COMPILE %s && %RUN | %CHECK %s

// SHR on unsigned BYTE must use logical shift (zero-fill), not arithmetic shift
FUNCTION main
VAR
    b : BYTE;
    s : SINT;
END_VAR
b := SHR(BYTE#251, SINT#1);

// CHECK: 125
printf('%d$N', b);

s := SHR(SINT#-4, SINT#1);

// CHECK: -2
printf('%d$N', s);
END_FUNCTION

(* ---- sizeof_arguments.st ---- *)
// RUN: %COMPILE %s && %RUN | %CHECK %s
//
// SIZEOF gives the same result for the implicit (positional) and the explicit (named) call form.

FUNCTION main
VAR
    arr : ARRAY[0..9] OF BYTE := [0, 1, 2, 3, 4, 5, 6, 7, 8, 9];
    a   : DINT;
    b   : DINT;
END_VAR

a := SIZEOF(arr);
b := SIZEOF(IN := arr);
// CHECK: SIZEOF=10 10
printf('SIZEOF=%d %d$N', a, b);
END_FUNCTION

(* ---- sub_arguments.st ---- *)
// RUN: %COMPILE %s && %RUN | %CHECK %s
//
// SUB gives the same result for the implicit (positional) and the explicit (named) call form, in
// declaration order and reordered. A call may also mix both forms: a named argument claims the slot
// its name declares, and the positional arguments fill the remaining slots in the order they are
// written.

FUNCTION main
VAR
    x   : DINT  := 9;
    y   : DINT  := 7331;
    lr  : LREAL := 1.5;
    lrr : LREAL;
    a   : DINT;
    b   : DINT;
    c   : DINT;
END_VAR

a := SUB(y, x);
b := SUB(IN1 := y, IN2 := x);
c := SUB(IN2 := x, IN1 := y);
// CHECK: SUB=7322 7322 7322
printf('SUB=%d %d %d$N', a, b, c);

// named argument before the positional one, IN1 is filled by y
a := SUB(IN2 := x, y);
// CHECK: SUB-named-first=7322
printf('SUB-named-first=%d$N', a);

// arguments of a different type
lrr := SUB(lr, 1);
// CHECK: SUB-mixed-types=0.5
printf('SUB-mixed-types=%.1f$N', lrr);
lrr := SUB(IN1 := lr, IN2 := 1);
// CHECK: SUB-mixed-types-named=0.5
printf('SUB-mixed-types-named=%.1f$N', lrr);

// parenthesized arguments
lrr := SUB((lr), 1);
// CHECK: SUB-paren=0.5
printf('SUB-paren=%.1f$N', lrr);
lrr := SUB(IN1 := (lr), IN2 := 1);
// CHECK: SUB-paren-named=0.5
printf('SUB-paren-named=%.1f$N', lrr);
END_FUNCTION

(* ---- upper_bound_arguments.st ---- *)
// RUN: %COMPILE %s && %RUN | %CHECK %s
//
// UPPER_BOUND gives the same result for the implicit (positional) and the explicit (named) call form,
// in declaration order and reordered.

FUNCTION main
VAR
    arr : ARRAY[0..9] OF BYTE := [0, 1, 2, 3, 4, 5, 6, 7, 8, 9];
END_VAR

bounds(arr);
END_FUNCTION

FUNCTION bounds : DINT
VAR_IN_OUT
    vla : ARRAY[*] OF BYTE;
END_VAR
VAR
    dim : DINT := 1;
    a   : DINT;
    b   : DINT;
    c   : DINT;
END_VAR

a := UPPER_BOUND(vla, dim);
b := UPPER_BOUND(ARR := vla, DIM := dim);
c := UPPER_BOUND(DIM := dim, ARR := vla);
// CHECK: UPPER_BOUND=9 9 9
printf('UPPER_BOUND=%d %d %d$N', a, b, c);
END_FUNCTION

(* ---- xor_arguments.st ---- *)
// RUN: %COMPILE %s && %RUN | %CHECK %s
//
// XOR declares a single variadic parameter. A variadic parameter cannot be named, thus XOR has an
// implicit (positional) call form only. The form is extensible. XOR gives the same result as the
// `XOR` operator, for BOOL values as well as for bit and integer values.

FUNCTION main
VAR
    t : BOOL := TRUE;
    f : BOOL := FALSE;
    x : BYTE := 16#F0;
    y : BYTE := 16#3C;
    z : BYTE := 16#01;
    i : DINT := 12;
    j : DINT := 10;
    a : BOOL;
    b : BOOL;
    c : BYTE;
    d : BYTE;
    e : DINT;
END_VAR

a := XOR(t, f);
b := XOR(t, f, t);
// CHECK: XOR=1 0 1 0
printf('XOR=%u %u %u %u$N', a, b, t XOR f, t XOR f XOR t);

c := XOR(x, y);
d := XOR(x, y, z);
e := XOR(i, j);
// CHECK: XOR-bits=204 205 6
printf('XOR-bits=%u %u %d$N', c, d, e);
// CHECK: XOR-bits-operator=204 205 6
printf('XOR-bits-operator=%u %u %d$N', x XOR y, x XOR y XOR z, i XOR j);
END_FUNCTION
